Staubli VAL3: main.pgx

program main()
begin
  close(tCurrentTool)
  pPointRs.config.shoulder = lefty
  pPointRs2.config.shoulder = lefty
  mCurrentSpeed.tvel = 100.00
  mCurrentSpeed.blend = joint
  mCurrentSpeed.reach = 0.010
  mCurrentSpeed.leave = 0.010
  call MoveJoint(30.00000,25.00000,80.00000,-45.00000)
  call MoveJoint(10.00000,-20.00000,50.00000,30.00000)
  call MoveJoint(30.00000,25.00000,80.00000,-45.00000)
  call MoveJoint(10.00000,-20.00000,50.00000,30.00000)
  call MoveJoint(30.00000,25.00000,80.00000,-45.00000)
  call MoveJoint(10.00000,-20.00000,50.00000,30.00000)

end
